RESOURCE RES0 : EMB_RES_ECO
  FBS
    RobotsStation : RoboCat;
    CapDist : CapDistributionCAT;
    APP_INIT : EVENTCHAINHEAD(NAME := 'APP_INIT');
  END_FBS
  EVENT_CONNECTIONS
    RobotsStation.A39BFC97654CAFF3 TO CapDist.E4C6FDAF265EC198;
    START.COLD TO APP_INIT.INIT;
    START.WARM TO APP_INIT.INIT;
    APP_INIT.INITO TO APP_INIT.TRIGGER;
    START.COLD TO RobotsStation.AEFC9DC06D949578;
    START.WARM TO RobotsStation.AEFC9DC06D949578;
  END_CONNECTIONS
END_RESOURCE
